(* PLC project PR_IRVisionCheckSeq_Soft2.0 1_workflow_93eeda_PLC, SiemensToBackhoff Siemens TIA Portal → Beckhoff TwinCAT PLCopen Converter 2.2 *)
(* stored: creationDateTime 2026-10-12T09:24:53.804929, modificationDateTime 2026-10-12T09:24:53.804929 *)

FUNCTION_BLOCK PR_IRVisionCheckSeq_Soft2.0 1_workflow_93eeda
VAR_INPUT
	iAutoRunning : BOOL;
	iFaultReset : BOOL;
	iIRMesaureProbeDown : BOOL;
	iIRMesaureProbeUp : BOOL;
	iIndexCylHome : BOOL;
	iIndexProbeOut : BOOL;
	iInspectionOver : BOOL;
	iManualEntryConfirm : BOOL;
	iMesauringOver : BOOL;
	iProbeCylHome : BOOL;
	iRFIDReadError : BOOL;
	iRFIDReadOver : BOOL;
	iReject : BOOL;
	iReset_fault : BOOL;
	iRetry : BOOL;
	iRetryCount : INT;
	iSstMode : BOOL;
	iSstPB : BOOL;
	iStartFrmFibroseq : BOOL;
END_VAR
VAR_OUTPUT
	qCameraLight : BOOL;
	qError : ARRAY[0..9] OF BOOL;
	qIRProbeDown : BOOL;
	qIRProbeUp : BOOL;
	qIRVisionCheckOver : BOOL;
	qIndexProbeIn : BOOL;
	qIndexProbeOut : BOOL;
	qMessage : ARRAY[0..9] OF BOOL;
END_VAR
VAR
	c20_ChkRecoveryStatus_T1 : BOOL;
	c20_ChkRecoveryStatus_T2 : BOOL;
	c20_ChkRecoveryStatus_T3 : BOOL;
	c20_ChkRecoveryStatus_T4 : BOOL;
	c22_WtRFIDReadOver_T1 : BOOL;
	c22_WtRFIDReadOver_T2 : BOOL;
	c23_ChkRetryCountOver_T1 : BOOL;
	c23_ChkRetryCountOver_T2 : BOOL;
	c24_WtOperatorDecisionRead_T1 : BOOL;
	c24_WtOperatorDecisionRead_T2 : BOOL;
	c25_ChkPartWorkable_T1 : BOOL;
	c25_ChkPartWorkable_T2 : BOOL;
	c91_WtRFIDWriteOver_T1 : BOOL;
	c91_WtRFIDWriteOver_T2 : BOOL;
	c92_ChkWriteRetryCountOver_T1 : BOOL;
	c92_ChkWriteRetryCountOver_T2 : BOOL;
	c93_WtOperatorDecisionWrite_T1 : BOOL;
	c93_WtOperatorDecisionWrite_T2 : BOOL;
	StateNo : INT;
	s100_WtStartLow : BOOL;
	s100_WtStartLow_T1 : BOOL;
	s10_WtStartFrmFibroSeq : BOOL;
	s10_WtStartFrmFibroSeq_T1 : BOOL;
	s1_WtResetRel : BOOL;
	s1_WtResetRel_T1 : BOOL;
	s20_ChkRecoveryStatus : BOOL;
	s20_ChkRecoveryStatus_T1 : BOOL;
	s20_ChkRecoveryStatus_T2 : BOOL;
	s20_ChkRecoveryStatus_T3 : BOOL;
	s20_ChkRecoveryStatus_T4 : BOOL;
	s21_WtProbeIndexCylHome : BOOL;
	s21_WtProbeIndexCylHome_T1 : BOOL;
	s22_WtRFIDReadOver : BOOL;
	s22_WtRFIDReadOver_T1 : BOOL;
	s22_WtRFIDReadOver_T2 : BOOL;
	s23_ChkRetryCountOver : BOOL;
	s23_ChkRetryCountOver_T1 : BOOL;
	s23_ChkRetryCountOver_T2 : BOOL;
	s24_WtOperatorDecisionRead : BOOL;
	s24_WtOperatorDecisionRead_T1 : BOOL;
	s24_WtOperatorDecisionRead_T2 : BOOL;
	s25_ChkPartWorkable : BOOL;
	s25_ChkPartWorkable_T1 : BOOL;
	s25_ChkPartWorkable_T2 : BOOL;
	s30_WtOperatorAck : BOOL;
	s30_WtOperatorAck_T1 : BOOL;
	s50_WtIRMeasureProbeAtTest : BOOL;
	s50_WtIRMeasureProbeAtTest_T1 : BOOL;
	s60_WtMeasurementOver : BOOL;
	s60_WtMeasurementOver_T1 : BOOL;
	s70_WtIRMeasureProbeUp : BOOL;
	s70_WtIRMeasureProbeUp_T1 : BOOL;
	s80_WtIndexingProbeOut : BOOL;
	s80_WtIndexingProbeOut_T1 : BOOL;
	s90_WtVisionInspectionOver : BOOL;
	s90_WtVisionInspectionOver_T1 : BOOL;
	s91_WtRFIDWriteOver : BOOL;
	s91_WtRFIDWriteOver_T1 : BOOL;
	s91_WtRFIDWriteOver_T2 : BOOL;
	s92_ChkWriteRetryCountOver : BOOL;
	s92_ChkWriteRetryCountOver_T1 : BOOL;
	s92_ChkWriteRetryCountOver_T2 : BOOL;
	s93_WtOperatorDecisionWrite : BOOL;
	s93_WtOperatorDecisionWrite_T1 : BOOL;
	s93_WtOperatorDecisionWrite_T2 : BOOL;
	s94_WtAllSystemAtHome : BOOL;
	s94_WtAllSystemAtHome_T1 : BOOL;
	sAbnormalStatus : BOOL;
	sIRInProgress : BOOL;
	sPartWorkable : BOOL;
	sRFReadRetryCount : INT;
	sRFWriteError : BOOL;
	sRFWriteOver : BOOL;
	sRFWriteRetryCount : INT;
	sSst : BOOL;
	sSstPulse : BOOL;
	sSstRise : R_TRIG;
	sStWtResetRel : BOOL;
	sStWtResetRel_T1 : BOOL;
	sTimeouTime : TON;
	sVisionInProgress : BOOL;
END_VAR
VAR_TEMP
	tOne : BOOL;
END_VAR
  VAR  (* added by the conversion: wires and edge detectors of the diagram *)
    _w24 : BOOL;
    _w26 : BOOL;
    _w39 : BOOL;
    _w41 : BOOL;
    _w42 : BOOL;
    _w55 : BOOL;
    _w58 : BOOL;
    _w59 : BOOL;
    _w112 : BOOL;
    _w115 : BOOL;
    _w116 : BOOL;
    _w117 : BOOL;
    _w118 : BOOL;
    _w119 : BOOL;
    _w132 : BOOL;
    _w134 : BOOL;
    _w135 : BOOL;
    _w153 : BOOL;
    _w155 : BOOL;
    _w156 : BOOL;
    _w186 : BOOL;
    _w190 : BOOL;
    _w191 : BOOL;
    _w192 : BOOL;
    _w228 : BOOL;
    _w230 : BOOL;
    _w231 : BOOL;
    _w232 : BOOL;
    _w257 : BOOL;
    _w259 : BOOL;
    _w260 : BOOL;
    _w261 : BOOL;
    _w289 : BOOL;
    _w292 : BOOL;
    _w293 : BOOL;
    _w294 : BOOL;
    _w307 : BOOL;
    _w309 : BOOL;
    _w310 : BOOL;
    _w327 : BOOL;
    _w330 : BOOL;
    _w331 : BOOL;
    _w356 : BOOL;
    _w358 : BOOL;
    _w359 : BOOL;
    _w376 : BOOL;
    _w378 : BOOL;
    _w379 : BOOL;
    _w396 : BOOL;
    _w399 : BOOL;
    _w400 : BOOL;
    _w437 : BOOL;
    _w442 : BOOL;
    _w443 : BOOL;
    _w444 : BOOL;
    _w480 : BOOL;
    _w482 : BOOL;
    _w483 : BOOL;
    _w484 : BOOL;
    _w509 : BOOL;
    _w511 : BOOL;
    _w512 : BOOL;
    _w513 : BOOL;
    _w531 : BOOL;
    _w535 : BOOL;
    _w536 : BOOL;
    _w554 : BOOL;
    _w556 : BOOL;
    _w557 : BOOL;
  END_VAR

(* LD diagram, written out as Structured Text *)
(* Network 1 *)
(* Create Single Step Pulse bit *)
(* Create Single Step bit *)
(* Transition for STATE Num:0 Reset Released *)
(* STATE Num:0 Reset Released *)
(* Transition for STATE Num:1 Wait For Reset Release *)
(* STATE Num:1 Wait For Reset Release *)
(* Transition for STATE Num:10 Wait For Start From Fibro Main Seq *)
(* STATE Num:10 Wait For Start From Fibro Main Seq *)
(* Actions for STATE Num:10 Wait For Start From Fibro Main Seq *)
(* Condition1 for STATE Num:20 Check Recovery Status *)
(* Condition2 for STATE Num:20 Check Recovery Status *)
(* Condition3 for STATE Num:20 Check Recovery Status *)
(* Condition4 for STATE Num:20 Check Recovery Status *)
(* Transition for STATE Num:20 Check Recovery Status *)
(* STATE Num:20 Check Recovery Status *)
(* Transition for STATE Num:30 Wait for Operator Ack *)
(* STATE Num:30 Wait for Operator Ack *)
(* Actions for STATE Num:30 Wait for Operator Ack *)
(* Transition for STATE Num:21 Wait For Probe and Index Cyl Home *)
(* STATE Num:21 Wait For Probe and Index Cyl Home *)
(* Actions for STATE Num:21 Wait For Probe and Index Cyl Home *)
(* Condition1 for STATE Num:22 Wait For RFID Read Over *)
(* Condition2 for STATE Num:22 Wait For RFID Read Over *)
(* Transition for STATE Num:22 Wait For RFID Read Over *)
(* STATE Num:22 Wait For RFID Read Over *)
(* Transition Actions T1 for STATE Num:22 Wait For RFID Read Over *)
(* Condition1 for STATE Num:23 Check Retry Count Over *)
(* Condition2 for STATE Num:23 Check Retry Count Over *)
(* Transition for STATE Num:23 Check Retry Count Over *)
(* STATE Num:23 Check Retry Count Over *)
(* Condition1 for STATE Num:24 Wait For Operator Decision_Read *)
(* Condition2 for STATE Num:24 Wait For Operator Decision_Read *)
(* Transition for STATE Num:24 Wait For Operator Decision_Read *)
(* STATE Num:24 Wait For Operator Decision_Read *)
(* Actions for STATE Num:24 Wait For Operator Decision_Read *)
(* Condition1 for STATE Num:25 Check Part is Workable *)
(* Condition2 for STATE Num:25 Check Part is Workable *)
(* Transition for STATE Num:25 Check Part is Workable *)
(* STATE Num:25 Check Part is Workable *)
(* Transition for STATE Num:50 Wait for IR Measure Probe At Test *)
(* STATE Num:50 Wait for IR Measure Probe At Test *)
(* Actions for STATE Num:50 Wait for IR Measure Probe At Test *)
(* Transition for STATE Num:60 Wait For Measurement Over *)
(* STATE Num:60 Wait For Measurement Over *)
(* Network 46 *)
(* Transition for STATE Num:70 Wait For IR Measure Probe Up *)
(* STATE Num:70 Wait For IR Measure Probe Up *)
(* Actions for STATE Num:70 Wait For IR Measure Probe Up *)
(* Transition for STATE Num:80 Wait For Indexing Probe Out *)
(* STATE Num:80 Wait For Indexing Probe Out *)
(* Actions for STATE Num:80 Wait For Indexing Probe Out *)
(* Transition for STATE Num:90 Wait For Vision Inspection Over *)
(* STATE Num:90 Wait For Vision Inspection Over *)
(* Network 55 *)
(* Condition1 for STATE Num:91 Wait for RFID Write Over *)
(* Condition2 for STATE Num:91 Wait for RFID Write Over *)
(* Transition for STATE Num:91 Wait for RFID Write Over *)
(* STATE Num:91 Wait for RFID Write Over *)
(* Network 60 *)
(* Condition1 for STATE Num:92 Check Write Retry Count Over *)
(* Condition2 for STATE Num:92 Check Write Retry Count Over *)
(* Transition for STATE Num:92 Check Write Retry Count Over *)
(* STATE Num:92 Check Write Retry Count Over *)
(* Condition1 for STATE Num:93 Wait For Operator Decision_Write *)
(* Condition2 for STATE Num:93 Wait For Operator Decision_Write *)
(* Transition for STATE Num:93 Wait For Operator Decision_Write *)
(* Network 68 *)
(* Actions for STATE Num:93 Wait For Operator Decision_Write *)
(* Transition for STATE Num:94 Wait for All System At Home *)
(* STATE Num:94 Wait for All System At Home *)
(* Actions for STATE Num:94 Wait for All System At Home *)
(* Transition for STATE Num:100 Wait For Start Low *)
(* STATE Num:100 Wait For Start Low *)
(* Network 75 *)
tOne := tOne OR NOT tOne;
sSstRise(CLK := iSstPB);
sSstPulse := sSstRise.Q;
sSst := iSstMode AND sSstPulse OR NOT iSstMode;
sStWtResetRel_T1 := sStWtResetRel AND iAutoRunning;
_w24 := sStWtResetRel;
_w26 := (_w24 OR NOT iAutoRunning) AND NOT sStWtResetRel_T1;
sStWtResetRel := _w26;
IF _w26 THEN StateNo := 0; END_IF;
s1_WtResetRel_T1 := s1_WtResetRel AND NOT sStWtResetRel AND sSst AND iAutoRunning;
_w39 := s1_WtResetRel;
_w41 := (_w39 OR sStWtResetRel_T1) AND NOT sStWtResetRel;
_w42 := _w41 AND NOT s1_WtResetRel_T1;
s1_WtResetRel := _w42;
IF _w42 THEN StateNo := 1; END_IF;
s10_WtStartFrmFibroSeq_T1 := s10_WtStartFrmFibroSeq AND NOT sStWtResetRel AND sSst AND iStartFrmFibroseq;
_w55 := s10_WtStartFrmFibroSeq;
_w58 := (_w55 OR s1_WtResetRel_T1 OR s100_WtStartLow_T1) AND NOT sStWtResetRel;
_w59 := _w58 AND NOT s10_WtStartFrmFibroSeq_T1;
s10_WtStartFrmFibroSeq := _w59;
IF _w59 THEN StateNo := 10; END_IF;
IF s10_WtStartFrmFibroSeq THEN sRFReadRetryCount := 0; END_IF;
IF s10_WtStartFrmFibroSeq THEN sRFWriteRetryCount := 0; END_IF;
c20_ChkRecoveryStatus_T1 := sAbnormalStatus;
c20_ChkRecoveryStatus_T2 := NOT sAbnormalStatus AND sVisionInProgress;
c20_ChkRecoveryStatus_T3 := NOT sAbnormalStatus AND NOT sVisionInProgress AND sIRInProgress;
c20_ChkRecoveryStatus_T4 := NOT sAbnormalStatus AND NOT sVisionInProgress AND NOT sIRInProgress;
s20_ChkRecoveryStatus_T1 := s20_ChkRecoveryStatus AND NOT sStWtResetRel AND sSst AND c20_ChkRecoveryStatus_T1;
s20_ChkRecoveryStatus_T2 := s20_ChkRecoveryStatus AND NOT sStWtResetRel AND sSst AND NOT s20_ChkRecoveryStatus_T1 AND c20_ChkRecoveryStatus_T2;
s20_ChkRecoveryStatus_T3 := s20_ChkRecoveryStatus AND NOT sStWtResetRel AND sSst AND NOT s20_ChkRecoveryStatus_T1 AND NOT s20_ChkRecoveryStatus_T2 AND c20_ChkRecoveryStatus_T3;
s20_ChkRecoveryStatus_T4 := s20_ChkRecoveryStatus AND NOT sStWtResetRel AND sSst AND NOT s20_ChkRecoveryStatus_T1 AND NOT s20_ChkRecoveryStatus_T2 AND NOT s20_ChkRecoveryStatus_T3 AND c20_ChkRecoveryStatus_T4;
_w112 := s20_ChkRecoveryStatus;
_w115 := (_w112 OR s10_WtStartFrmFibroSeq_T1 OR s30_WtOperatorAck_T1) AND NOT sStWtResetRel;
_w116 := _w115 AND NOT s20_ChkRecoveryStatus_T1;
_w117 := _w116 AND NOT s20_ChkRecoveryStatus_T2;
_w118 := _w117 AND NOT s20_ChkRecoveryStatus_T3;
_w119 := _w118 AND NOT s20_ChkRecoveryStatus_T4;
s20_ChkRecoveryStatus := _w119;
IF _w119 THEN StateNo := 20; END_IF;
s30_WtOperatorAck_T1 := s30_WtOperatorAck AND NOT sStWtResetRel AND sSst AND iFaultReset;
_w132 := s30_WtOperatorAck;
_w134 := (_w132 OR s20_ChkRecoveryStatus_T1) AND NOT sStWtResetRel;
_w135 := _w134 AND NOT s30_WtOperatorAck_T1;
s30_WtOperatorAck := _w135;
IF _w135 THEN StateNo := 30; END_IF;
qError[0] := s30_WtOperatorAck;
s21_WtProbeIndexCylHome_T1 := s21_WtProbeIndexCylHome AND NOT sStWtResetRel AND sSst AND iProbeCylHome AND iIndexCylHome;
_w153 := s21_WtProbeIndexCylHome;
_w155 := (_w153 OR s20_ChkRecoveryStatus_T4) AND NOT sStWtResetRel;
_w156 := _w155 AND NOT s21_WtProbeIndexCylHome_T1;
s21_WtProbeIndexCylHome := _w156;
IF _w156 THEN StateNo := 21; END_IF;
qIRProbeUp := s21_WtProbeIndexCylHome;
qIndexProbeIn := s21_WtProbeIndexCylHome;
c22_WtRFIDReadOver_T1 := iRFIDReadError;
c22_WtRFIDReadOver_T2 := NOT iRFIDReadError AND iRFIDReadOver;
s22_WtRFIDReadOver_T1 := s22_WtRFIDReadOver AND NOT sStWtResetRel AND sSst AND c22_WtRFIDReadOver_T1;
s22_WtRFIDReadOver_T2 := s22_WtRFIDReadOver AND NOT sStWtResetRel AND sSst AND NOT s22_WtRFIDReadOver_T1 AND c22_WtRFIDReadOver_T2;
_w186 := s22_WtRFIDReadOver;
_w190 := (_w186 OR s21_WtProbeIndexCylHome_T1 OR s23_ChkRetryCountOver_T2 OR s24_WtOperatorDecisionRead_T1) AND NOT sStWtResetRel;
_w191 := _w190 AND NOT s22_WtRFIDReadOver_T1;
_w192 := _w191 AND NOT s22_WtRFIDReadOver_T2;
s22_WtRFIDReadOver := _w192;
IF _w192 THEN StateNo := 22; END_IF;
IF s22_WtRFIDReadOver_T1 THEN sRFReadRetryCount := sRFReadRetryCount + 1; END_IF;
qMessage[0] := s22_WtRFIDReadOver;
c23_ChkRetryCountOver_T1 := sRFReadRetryCount > iRetryCount;
c23_ChkRetryCountOver_T2 := sRFReadRetryCount <= iRetryCount;
s23_ChkRetryCountOver_T1 := s23_ChkRetryCountOver AND NOT sStWtResetRel AND sSst AND c23_ChkRetryCountOver_T1;
s23_ChkRetryCountOver_T2 := s23_ChkRetryCountOver AND NOT sStWtResetRel AND sSst AND NOT s23_ChkRetryCountOver_T1 AND c23_ChkRetryCountOver_T2;
_w228 := s23_ChkRetryCountOver;
_w230 := (_w228 OR s22_WtRFIDReadOver_T1) AND NOT sStWtResetRel;
_w231 := _w230 AND NOT s23_ChkRetryCountOver_T1;
_w232 := _w231 AND NOT s23_ChkRetryCountOver_T2;
s23_ChkRetryCountOver := _w232;
IF _w232 THEN StateNo := 23; END_IF;
c24_WtOperatorDecisionRead_T1 := iRetry;
c24_WtOperatorDecisionRead_T2 := NOT iRetry AND iManualEntryConfirm;
s24_WtOperatorDecisionRead_T1 := s24_WtOperatorDecisionRead AND NOT sStWtResetRel AND sSst AND c24_WtOperatorDecisionRead_T1;
s24_WtOperatorDecisionRead_T2 := s24_WtOperatorDecisionRead AND NOT sStWtResetRel AND sSst AND NOT s24_WtOperatorDecisionRead_T1 AND c24_WtOperatorDecisionRead_T2;
_w257 := s24_WtOperatorDecisionRead;
_w259 := (_w257 OR s23_ChkRetryCountOver_T1) AND NOT sStWtResetRel;
_w260 := _w259 AND NOT s24_WtOperatorDecisionRead_T1;
_w261 := _w260 AND NOT s24_WtOperatorDecisionRead_T2;
s24_WtOperatorDecisionRead := _w261;
IF _w261 THEN StateNo := 24; END_IF;
qError[5] := s24_WtOperatorDecisionRead;
c25_ChkPartWorkable_T1 := NOT sPartWorkable;
c25_ChkPartWorkable_T2 := sPartWorkable;
s25_ChkPartWorkable_T1 := s25_ChkPartWorkable AND NOT sStWtResetRel AND sSst AND c25_ChkPartWorkable_T1;
s25_ChkPartWorkable_T2 := s25_ChkPartWorkable AND NOT sStWtResetRel AND sSst AND NOT s25_ChkPartWorkable_T1 AND c25_ChkPartWorkable_T2;
_w289 := s25_ChkPartWorkable;
_w292 := (_w289 OR s22_WtRFIDReadOver_T2 OR s24_WtOperatorDecisionRead_T2) AND NOT sStWtResetRel;
_w293 := _w292 AND NOT s25_ChkPartWorkable_T1;
_w294 := _w293 AND NOT s25_ChkPartWorkable_T2;
s25_ChkPartWorkable := _w294;
IF _w294 THEN StateNo := 25; END_IF;
s50_WtIRMeasureProbeAtTest_T1 := s50_WtIRMeasureProbeAtTest AND NOT sStWtResetRel AND sSst AND iIRMesaureProbeDown;
_w307 := s50_WtIRMeasureProbeAtTest;
_w309 := (_w307 OR s25_ChkPartWorkable_T2) AND NOT sStWtResetRel;
_w310 := _w309 AND NOT s50_WtIRMeasureProbeAtTest_T1;
s50_WtIRMeasureProbeAtTest := _w310;
IF _w310 THEN StateNo := 50; END_IF;
qIRProbeDown := s50_WtIRMeasureProbeAtTest;
s60_WtMeasurementOver_T1 := s60_WtMeasurementOver AND NOT sStWtResetRel AND sSst AND iMesauringOver;
_w327 := s60_WtMeasurementOver;
_w330 := (_w327 OR s50_WtIRMeasureProbeAtTest_T1 OR s20_ChkRecoveryStatus_T3) AND NOT sStWtResetRel;
_w331 := _w330 AND NOT s60_WtMeasurementOver_T1;
s60_WtMeasurementOver := _w331;
IF _w331 THEN StateNo := 60; END_IF;
sTimeouTime(IN := s60_WtMeasurementOver AND NOT iMesauringOver, PT := t#5s);
qError[1] := s60_WtMeasurementOver AND NOT iMesauringOver AND sTimeouTime.Q OR qError[1] AND NOT iFaultReset;
s70_WtIRMeasureProbeUp_T1 := s70_WtIRMeasureProbeUp AND NOT sStWtResetRel AND sSst AND iIRMesaureProbeUp;
_w356 := s70_WtIRMeasureProbeUp;
_w358 := (_w356 OR s60_WtMeasurementOver_T1) AND NOT sStWtResetRel;
_w359 := _w358 AND NOT s70_WtIRMeasureProbeUp_T1;
s70_WtIRMeasureProbeUp := _w359;
IF _w359 THEN StateNo := 70; END_IF;
qIRProbeUp := s70_WtIRMeasureProbeUp;
s80_WtIndexingProbeOut_T1 := s80_WtIndexingProbeOut AND NOT sStWtResetRel AND sSst AND iIndexProbeOut;
_w376 := s80_WtIndexingProbeOut;
_w378 := (_w376 OR s70_WtIRMeasureProbeUp_T1) AND NOT sStWtResetRel;
_w379 := _w378 AND NOT s80_WtIndexingProbeOut_T1;
s80_WtIndexingProbeOut := _w379;
IF _w379 THEN StateNo := 80; END_IF;
qIndexProbeOut := s80_WtIndexingProbeOut;
s90_WtVisionInspectionOver_T1 := s90_WtVisionInspectionOver AND NOT sStWtResetRel AND sSst AND iInspectionOver;
_w396 := s90_WtVisionInspectionOver;
_w399 := (_w396 OR s80_WtIndexingProbeOut_T1 OR s20_ChkRecoveryStatus_T2) AND NOT sStWtResetRel;
_w400 := _w399 AND NOT s90_WtVisionInspectionOver_T1;
s90_WtVisionInspectionOver := _w400;
IF _w400 THEN StateNo := 90; END_IF;
sTimeouTime(IN := s90_WtVisionInspectionOver AND NOT iInspectionOver, PT := t#5s);
qError[2] := s90_WtVisionInspectionOver AND NOT iInspectionOver AND sTimeouTime.Q OR qError[2] AND NOT iFaultReset;
c91_WtRFIDWriteOver_T1 := sRFWriteError;
c91_WtRFIDWriteOver_T2 := NOT sRFWriteError AND sRFWriteOver;
s91_WtRFIDWriteOver_T1 := s91_WtRFIDWriteOver AND NOT sStWtResetRel AND sSst AND c91_WtRFIDWriteOver_T1;
s91_WtRFIDWriteOver_T2 := s91_WtRFIDWriteOver AND NOT sStWtResetRel AND sSst AND NOT s91_WtRFIDWriteOver_T1 AND c91_WtRFIDWriteOver_T2;
_w437 := s91_WtRFIDWriteOver;
_w442 := (_w437 OR s90_WtVisionInspectionOver_T1 OR s25_ChkPartWorkable_T1 OR s92_ChkWriteRetryCountOver_T2 OR s93_WtOperatorDecisionWrite_T2) AND NOT sStWtResetRel;
_w443 := _w442 AND NOT s91_WtRFIDWriteOver_T1;
_w444 := _w443 AND NOT s91_WtRFIDWriteOver_T2;
s91_WtRFIDWriteOver := _w444;
IF _w444 THEN StateNo := 91; END_IF;
qMessage[1] := s91_WtRFIDWriteOver;
IF s91_WtRFIDWriteOver_T1 THEN sRFWriteRetryCount := sRFWriteRetryCount + 1; END_IF;
c92_ChkWriteRetryCountOver_T1 := sRFWriteRetryCount > iRetryCount;
c92_ChkWriteRetryCountOver_T2 := sRFWriteRetryCount <= iRetryCount;
s92_ChkWriteRetryCountOver_T1 := s92_ChkWriteRetryCountOver AND NOT sStWtResetRel AND sSst AND c92_ChkWriteRetryCountOver_T1;
s92_ChkWriteRetryCountOver_T2 := s92_ChkWriteRetryCountOver AND NOT sStWtResetRel AND sSst AND NOT s92_ChkWriteRetryCountOver_T1 AND c92_ChkWriteRetryCountOver_T2;
_w480 := s92_ChkWriteRetryCountOver;
_w482 := (_w480 OR s91_WtRFIDWriteOver_T1) AND NOT sStWtResetRel;
_w483 := _w482 AND NOT s92_ChkWriteRetryCountOver_T1;
_w484 := _w483 AND NOT s92_ChkWriteRetryCountOver_T2;
s92_ChkWriteRetryCountOver := _w484;
IF _w484 THEN StateNo := 92; END_IF;
c93_WtOperatorDecisionWrite_T1 := iReject;
c93_WtOperatorDecisionWrite_T2 := NOT iReject AND iRetry;
s93_WtOperatorDecisionWrite_T1 := s93_WtOperatorDecisionWrite AND NOT sStWtResetRel AND sSst AND c93_WtOperatorDecisionWrite_T1;
s93_WtOperatorDecisionWrite_T2 := s93_WtOperatorDecisionWrite AND NOT sStWtResetRel AND sSst AND NOT s93_WtOperatorDecisionWrite_T1 AND c93_WtOperatorDecisionWrite_T2;
_w509 := s93_WtOperatorDecisionWrite;
_w511 := (_w509 OR s92_ChkWriteRetryCountOver_T1) AND NOT sStWtResetRel;
_w512 := _w511 AND NOT s93_WtOperatorDecisionWrite_T1;
_w513 := _w512 AND NOT s93_WtOperatorDecisionWrite_T2;
s93_WtOperatorDecisionWrite := _w513;
IF _w513 THEN StateNo := 93; END_IF;
qError[6] := s93_WtOperatorDecisionWrite;
s94_WtAllSystemAtHome_T1 := s94_WtAllSystemAtHome AND NOT sStWtResetRel AND sSst AND iProbeCylHome AND iIndexCylHome;
_w531 := s94_WtAllSystemAtHome;
_w535 := (_w531 OR s92_ChkWriteRetryCountOver_T1 OR s93_WtOperatorDecisionWrite_T1 OR s91_WtRFIDWriteOver_T2) AND NOT sStWtResetRel;
_w536 := _w535 AND NOT s94_WtAllSystemAtHome_T1;
s94_WtAllSystemAtHome := _w536;
IF _w536 THEN StateNo := 94; END_IF;
qIRProbeUp := s94_WtAllSystemAtHome;
qIndexProbeIn := s94_WtAllSystemAtHome;
s100_WtStartLow_T1 := s100_WtStartLow AND NOT sStWtResetRel AND sSst AND NOT iStartFrmFibroseq;
_w554 := s100_WtStartLow;
_w556 := (_w554 OR s94_WtAllSystemAtHome_T1) AND NOT sStWtResetRel;
_w557 := _w556 AND NOT s100_WtStartLow_T1;
s100_WtStartLow := _w557;
IF _w557 THEN StateNo := 100; END_IF;
IF iStartFrmFibroseq THEN sIRInProgress := FALSE; END_IF;
IF iStartFrmFibroseq THEN sVisionInProgress := FALSE; END_IF;
IF s100_WtStartLow THEN qIRVisionCheckOver := TRUE; END_IF;
IF iStartFrmFibroseq THEN sRFReadRetryCount := 0; END_IF;
IF iStartFrmFibroseq THEN sRFWriteRetryCount := 0; END_IF;
END_FUNCTION_BLOCK
